(* IEC 61131-3 sources: 2026_Projet_YGO_ExcavatriceDragage/ARCHIVES/Code/CFC_STAGING_RECOVERED/CODE/COMMUN, 2 files *)

(* ---- ST_ResetCommand.st ---- *)
(* ═══════════════════════════════════════════════════════════════
   🔘 ST_ResetCommand — Commande Reset publique amont
   ───────────────────────────────────────────────────────────────
   🎯 Niveau continu issu de l'IHM. Chaque consommateur porte son
      propre détecteur de front : ce contrat ne mémorise aucun état.
   🛡️ Un Reset ne réarme jamais sans action consciente ultérieure.
   ═══════════════════════════════════════════════════════════════ *)
TYPE ST_ResetCommand :
STRUCT
    CmdReset : BOOL;  (* TRUE = au moins une demande Reset IHM présente *)
END_STRUCT
END_TYPE

(* ---- FB_ResetAggregation.st ---- *)
(* ═══════════════════════════════════════════════════════════════
   🔘 FB_ResetAggregation — Producteur unique du niveau Reset IHM
   ───────────────────────────────────────────────────────────────
   📄 Contrat : ST_ResetCommand
   🛡️ Agrège uniquement les quatre boutons existants. Il ne détecte
      pas de front et ne réarme rien : les consommateurs conservent
      leur R_TRIG local, conformément à la règle Reset = front.
   ═══════════════════════════════════════════════════════════════ *)
FUNCTION_BLOCK FB_ResetAggregation
VAR_INPUT
    BtnFaultReset : BOOL;
    BtnResetM1 : BOOL;
    BtnResetM2 : BOOL;
    BtnResetBucket : BOOL;
END_VAR
VAR_OUTPUT
    Cmd : ST_ResetCommand;
END_VAR

Cmd.CmdReset := BtnFaultReset OR BtnResetM1 OR BtnResetM2 OR BtnResetBucket;
